FUNCTION_BLOCK FB_MovingAverage_Test EXTENDS TcUnit.FB_TestSuite

calculationShouldBeReadyWhenTimePassed();
calculationShouldNotBeReadyBeforeTimePassed();
movingAverageOfThreePlusTwoPlusOneShouldBeTwo();
resetMethodCallShouldResetValue();
theValueShouldBe40AfterTwoSeconds();
valueShouldBe0BeforeWindowPassedIfPreReadyNotIncluded();

METHOD calculationShouldBeReadyWhenTimePassed : BOOL
VAR
	movingAverage : FB_MovingAverage;
END_VAR

TEST('calculationShouldBeReadyWhenTimePassed');
movingAverage.startCalculation(TRUE,0, 3,1, T#3S, FALSE);
AssertEquals_BOOL(Expected := TRUE, Actual :=  movingAverage.ready, Message := 'Moving average calculation not ready after time passed');
TEST_FINISHED();
END_METHOD

METHOD calculationShouldNotBeReadyBeforeTimePassed : BOOL
VAR
	movingAverage : FB_MovingAverage;
END_VAR

TEST('calculationShouldNotBeReadyBeforeTimePassed');
movingAverage.startCalculation(TRUE, 0, 1,1, T#0S, FALSE);
AssertEquals_BOOL(Expected := FALSE, Actual :=  movingAverage.ready, Message := 'Moving average calculation ready before time passed');
TEST_FINISHED();
END_METHOD

METHOD movingAverageOfThreePlusTwoPlusOneShouldBeTwo
VAR
	movingAverage : FB_MovingAverage;
END_VAR

TEST('movingAverageOfThreePlusTwoPlusOneShouldBeTwo');
movingAverage.startCalculation(TRUE, 3, 3, 1, T#1S, FALSE);
movingAverage.startCalculation(TRUE, 2, 3, 1, T#1S, FALSE);
movingAverage.startCalculation(TRUE, 1, 3, 1, T#1S, FALSE);
movingAverage.startCalculation(TRUE, 0, 3, 1, T#1S, FALSE);
AssertEquals_REAL(Expected := 2, Actual := movingAverage.value, 0, Message := 'Moving average calculation not equal to two!');
TEST_FINISHED();
END_METHOD

METHOD resetMethodCallShouldResetValue
VAR
	movingAverage : FB_MovingAverage;
END_VAR

TEST('resetMethodCallShouldResetValue');
movingAverage.startCalculation(start := TRUE, measurement := 50, intervalS := 1, windowS := 3, dtime := T#3S, excludeUntilReady := FALSE);
movingAverage.reset();
AssertEquals_REAL(0, movingAverage.value, 0, 'Reset did not reset value!'); 
TEST_FINISHED();
END_METHOD

METHOD theValueShouldBe40AfterTwoSeconds
VAR
	movingAverage : FB_MovingAverage;
END_VAR
TEST('theValueShouldBe40AfterTwoSeconds');
movingAverage.startCalculation(start := TRUE, measurement := 40, intervalS := 1, windowS := 3, dtime := T#1S, excludeUntilReady := FALSE);
movingAverage.startCalculation(start := TRUE, measurement := 40, intervalS := 1, windowS := 3, dtime := T#1S, excludeUntilReady := FALSE);
AssertEquals_REAL(40, movingAverage.value, 0, 'Value not 40 after two seconds'); 
TEST_FINISHED();
END_METHOD

METHOD valueShouldBe0BeforeWindowPassedIfPreReadyNotIncluded
VAR
	movingAverage : FB_MovingAverage;
END_VAR

TEST('valueShouldBe0BeforeWindowPassedIfPreReadyNotIncluded');
movingAverage.startCalculation(start := TRUE, measurement := 40, intervalS := 1, windowS := 3, dtime := T#1S, excludeUntilReady := TRUE);
movingAverage.startCalculation(start := TRUE, measurement := 40, intervalS := 1, windowS := 3, dtime := T#1S, excludeUntilReady := TRUE);
AssertEquals_REAL(0, movingAverage.value, 0, 'Value not 0 before window passed when exclude values before first window checked'); 
TEST_FINISHED();
END_METHOD

END_FUNCTION_BLOCK

(* stored: Version 1.1.0.1, ProductVersion 3.1.4024.9
   POU FB_MovingAverage_Test: Id {2f19abed-84d4-48fe-930a-61fce21e2a0f}, SpecialFunc None
   Method calculationShouldBeReadyWhenTimePassed: Id {191212e6-4fc8-4265-bb95-62915115aacc}
   Method calculationShouldNotBeReadyBeforeTimePassed: Id {0f72b63f-fd9f-47d6-819b-ef24d985cb05}
   Method movingAverageOfThreePlusTwoPlusOneShouldBeTwo: Id {b9507e38-3aba-4d26-bc53-9f4ae707268f}
   Method resetMethodCallShouldResetValue: Id {a712c06f-d26e-4670-bdb3-b535903dbd74}
   Method theValueShouldBe40AfterTwoSeconds: Id {6d1812bd-834f-47d8-8609-a5c345ed96bf}
   Method valueShouldBe0BeforeWindowPassedIfPreReadyNotIncluded: Id {c81eda91-7c4d-4094-bd68-f8838112ac65} *)
